// TIA Portal V19 export
DATA_BLOCK "ALL_AI_DB"   // DB12
// stored: InstanceOfName ALL_AI, InstanceOfType FB
"ALL_AI"
   // VAR
   //    AI_TT01 { S7_SetPoint := 'True'} : "AI";
   //    AI_TT02 { S7_SetPoint := 'True'} : "AI";
   //    AI_TT03 { S7_SetPoint := 'True'} : "AI";
   //    AI_CHS_TT01 { S7_SetPoint := 'True'} : "AI";
   //    AI_CHS_TT02 { S7_SetPoint := 'True'} : "AI";
   //    AI_CHS_TT03 { S7_SetPoint := 'True'} : "AI";
   //    AI_CHS_TT04 { S7_SetPoint := 'True'} : "AI";
   //    AI_CHS_MGLT { S7_SetPoint := 'True'} : "AI";
   //    AI_R2_TT01 { S7_SetPoint := 'True'} : "AI";
   //    AI_R2_TT02 { S7_SetPoint := 'True'} : "AI";
   //    AI_R2_TT03 { S7_SetPoint := 'True'} : "AI";
   //    AI_R3_TT01 { S7_SetPoint := 'True'} : "AI";
   //    AI_R3_TT02 { S7_SetPoint := 'True'} : "AI";
   //    AI_R3_TT03 { S7_SetPoint := 'True'} : "AI";
   //    AI_R4_TT03 { S7_SetPoint := 'True'} : "AI";
   //    AI_R4_TT02 { S7_SetPoint := 'True'} : "AI";
   //    AI_R4_TT01 { S7_SetPoint := 'True'} : "AI";
   //    AI_R5_TT01 { S7_SetPoint := 'True'} : "AI";
   //    AI_R5_TT02 { S7_SetPoint := 'True'} : "AI";
   //    AI_R5_TT03 { S7_SetPoint := 'True'} : "AI";
   //    AI_R6_TT01 { S7_SetPoint := 'True'} : "AI";
   //    AI_R6_TT02 { S7_SetPoint := 'True'} : "AI";
   //    AI_R6_TT03 { S7_SetPoint := 'True'} : "AI";
   //    AI_R7_TT01 { S7_SetPoint := 'True'} : "AI";
   //    AI_R7_TT02 { S7_SetPoint := 'True'} : "AI";
   //    AI_R8_TT03 { S7_SetPoint := 'True'} : "AI";
   //    AI_R7_TT03 { S7_SetPoint := 'True'} : "AI";
   //    AI_R8_TT01 { S7_SetPoint := 'True'} : "AI";
   //    AI_R8_TT02 { S7_SetPoint := 'True'} : "AI";
   //    AI_R9_TT01 { S7_SetPoint := 'True'} : "AI";
   //    AI_R9_TT02 { S7_SetPoint := 'True'} : "AI";
   //    AI_R9_TT03 { S7_SetPoint := 'True'} : "AI";
   //    AI_R10_TT01 { S7_SetPoint := 'True'} : "AI";
   //    AI_R10_TT02 { S7_SetPoint := 'True'} : "AI";
   //    AI_R10_TT03 { S7_SetPoint := 'True'} : "AI";
   //    AI_R11_TT01 { S7_SetPoint := 'True'} : "AI";
   //    AI_R11_TT02 { S7_SetPoint := 'True'} : "AI";
   //    AI_R11_TT03 { S7_SetPoint := 'True'} : "AI";
   //    AI_R12_TT01 { S7_SetPoint := 'True'} : "AI";
   //    AI_R12_TT02 { S7_SetPoint := 'True'} : "AI";
   //    AI_R12_TT03 { S7_SetPoint := 'True'} : "AI";
   //    AI_R13_TT01 { S7_SetPoint := 'True'} : "AI";
   //    AI_R13_TT02 { S7_SetPoint := 'True'} : "AI";
   //    AI_R13_TT03 { S7_SetPoint := 'True'} : "AI";
   //    AI_R14_TT01 { S7_SetPoint := 'True'} : "AI";
   //    AI_R14_TT02 { S7_SetPoint := 'True'} : "AI";
   //    AI_R14_TT03 { S7_SetPoint := 'True'} : "AI";
   //    AI_R15_TT01 { S7_SetPoint := 'True'} : "AI";
   //    AI_R15_TT02 { S7_SetPoint := 'True'} : "AI";
   //    AI_R15_TT03 { S7_SetPoint := 'True'} : "AI";
   //    AI_R16_TT01 { S7_SetPoint := 'True'} : "AI";
   //    AI_R16_TT02 { S7_SetPoint := 'True'} : "AI";
   //    AI_R16_TT03 { S7_SetPoint := 'True'} : "AI";
   //    AI_R17_TT01 { S7_SetPoint := 'True'} : "AI";
   //    AI_R17_TT02 { S7_SetPoint := 'True'} : "AI";
   //    AI_R17_TT03 { S7_SetPoint := 'True'} : "AI";
   //    AI_R18_TT01 { S7_SetPoint := 'True'} : "AI";
   //    AI_R18_TT02 { S7_SetPoint := 'True'} : "AI";
   //    AI_R18_TT03 { S7_SetPoint := 'True'} : "AI";
   //    AI_CHS_PT { S7_SetPoint := 'True'} : "AI";
   //    AI_SMHS_TT01 { S7_SetPoint := 'True'} : "AI";
   //    AI_SMHS_TT02 { S7_SetPoint := 'True'} : "AI";
   //    AI_SMHS_TT03 { S7_SetPoint := 'True'} : "AI";
   //    AI_SMHS_TT04 { S7_SetPoint := 'True'} : "AI";
   //    AI_NMHS_TT01 { S7_SetPoint := 'True'} : "AI";
   //    AI_NMHS_TT02 { S7_SetPoint := 'True'} : "AI";
   //    AI_NMHS_TT03 { S7_SetPoint := 'True'} : "AI";
   //    AI_NMHS_TT04 { S7_SetPoint := 'True'} : "AI";
   //    AI_SMHS_PT01 { S7_SetPoint := 'True'} : "PT_AI";
   //    AI_SMHS_PT02 { S7_SetPoint := 'True'} : "PT_AI";
   //    AI_SMHS_PT03 { S7_SetPoint := 'True'} : "PT_AI";
   //    AI_SMHS_PT04 { S7_SetPoint := 'True'} : "PT_AI";
   //    AI_NMHS_PT04 { S7_SetPoint := 'True'} : "PT_AI";
   //    AI_NMHS_PT01 { S7_SetPoint := 'True'} : "PT_AI";
   //    AI_NMHS_PT02 { S7_SetPoint := 'True'} : "PT_AI";
   //    AI_NMHS_PT03 { S7_SetPoint := 'True'} : "PT_AI";
   //    AI_CS_TT01 { S7_SetPoint := 'True'} : "AI";
   //    AI_CS_TT02 { S7_SetPoint := 'True'} : "AI";
   //    AI_CS_TT03 { S7_SetPoint := 'True'} : "AI";
   //    AI_CS_TT04 { S7_SetPoint := 'True'} : "AI";
   //    AI_CS_MGLT { S7_SetPoint := 'True'} : "AI";
   //    AI_UCHS_TT01 { S7_SetPoint := 'True'} : "AI";
   //    AI_UCHS_TT02 { S7_SetPoint := 'True'} : "AI";
   //    AI_UCHS_TT03 { S7_SetPoint := 'True'} : "AI";
   //    AI_UCHS_TT04 { S7_SetPoint := 'True'} : "AI";
   //    AI_UCHS_MGLT { S7_SetPoint := 'True'} : "AI";
   //    AI_HS_TT01 { S7_SetPoint := 'True'} : "AI";
   //    AI_HS_TT02 { S7_SetPoint := 'True'} : "AI";
   //    AI_HS_TT03 { S7_SetPoint := 'True'} : "AI";
   //    AI_HS_MGLT { S7_SetPoint := 'True'} : "AI";
   //    "AI_A/SCRB_001_PH01" { S7_SetPoint := 'True'} : "AI";
   //    "AI_AI_A/SCRB_002_PH01" { S7_SetPoint := 'True'} : "AI";
   //    "AI_A/VP_01_APT01" { S7_SetPoint := 'True'} : "AI";
   //    "AI_A/VP_02_APT01" { S7_SetPoint := 'True'} : "AI";
   //    "AI_A/ANFD_001_APT01" { S7_SetPoint := 'True'} : "AI";
   //    "AI_A/ANFD_002_APT01" { S7_SetPoint := 'True'} : "AI";
   //    "AI_A/ANFD_003_APT01" { S7_SetPoint := 'True'} : "AI";
   //    AI_HS_TT9 { S7_SetPoint := 'True'} : "AI";
   //    "A/ANFD_001_TT01" { S7_SetPoint := 'True'} : "AI";
   //    "A/ANFD_002_TT01" { S7_SetPoint := 'True'} : "AI";
   //    "A/ANFD_003_TT01" { S7_SetPoint := 'True'} : "AI";
   //    "A/ANFD_004_TT01" { S7_SetPoint := 'True'} : "AI";
   //    AI_RCVD_001_APT01 { S7_SetPoint := 'True'} : "AI";
   //    AI_RCVD_002_APT01 { S7_SetPoint := 'True'} : "AI";
   //    AI_RCVD_001_TT01 { S7_SetPoint := 'True'} : "AI";
   //    AI_RCVD_002_TT01 { S7_SetPoint := 'True'} : "AI";
   //    "AI_A/VTD_001_APT01" { S7_SetPoint := 'True'} : "AI";
   //    "AI_A/VTD_002_APT01" { S7_SetPoint := 'True'} : "AI";
   //    "AI_A/VTD_001_TT01" { S7_SetPoint := 'True'} : "AI";
   //    "AI_A/VTD_002_TT01" { S7_SetPoint := 'True'} : "AI";
   //    "AI_A/TD_001_TT01" { S7_SetPoint := 'True'} : "AI";
   //    "AI_A/TD_002_TT01" { S7_SetPoint := 'True'} : "AI";
   //    DRIVE_RPM { S7_SetPoint := 'True'} : "DRIVE_RPM";
   // END_VAR
BEGIN
END_DATA_BLOCK
